Fanuc KAREL source: KB00157.KL

PROGRAM KB00157
%NOLOCKGROUP
%ENVIRONMENT MULTI
VAR
  P1: INTEGER
  RESULT: INTEGER
BEGIN
  P1 = 1
  RESULT = SEMA_COUNT(P1)
END KB00157
